(* IEC 61131-3 sources: virtual-bottling-plant/plc/src/process, 4 files *)

(* ---- FB_MixBatch.st ---- *)
(* T-101 batch sequence (PLC-03, ISA-88 phases): Fill (dose water, concentrate, sugar by
   flow totals), Mix, Transfer to T-301 through P-201. A recipe with another product first
   drains T-101 and T-301, then runs CIP. There is no time-of-day window: a new batch starts
   whenever T-101 is empty. One mix tank only (decision P2, see l1-plc.md). *)
FUNCTION_BLOCK FB_MixBatch
  VAR_INPUT
    Recipe : ST_Recipe;
    WaterFlow : REAL;        (* FT101, L/min *)
    ConcFlow : REAL;         (* FT102 *)
    SugarFlow : REAL;        (* FT103 *)
    Brix : REAL;             (* AT101 *)
    TankEmpty : BOOL;        (* LSL101 *)
    BufferLevel : REAL;      (* LT301, % *)
    CipDone : BOOL;
    NowMs : UDINT;
    DtS : REAL;
  END_VAR
  VAR_OUTPUT
    WaterValve : BOOL;
    ConcValve : BOOL;
    SugarValve : BOOL;
    Agitator : BOOL;
    TransferPump : BOOL;
    TankDrain : BOOL;
    BufferDrain : BOOL;
    CipRun : BOOL;
    ConcSelect : REAL;       (* product code to the concentrate feed selector *)
    Status : ST_T101Status;
    BrixAlarm : BOOL;
  END_VAR
  VAR
    MixTimer : FB_SimTon;
    NotEmptyInIdle : FB_SimTon;
    TargetWater : REAL;
    TargetConc : REAL;
    TargetSugar : REAL;
    DosedWater : REAL;
    DosedConc : REAL;
    DosedSugar : REAL;
    ConcBrix : REAL;
    PumpOn : BOOL;
  END_VAR
  VAR CONSTANT
    BATCH_L : REAL := 5000.0;
    SUGAR_SYRUP_BRIX : REAL := 67.0;
    MIX_MS : UDINT := 900000;        (* 15 min *)
    BUFFER_PUMP_ON : REAL := 90.0;   (* % T-301 *)
    BUFFER_PUMP_OFF : REAL := 98.0;
    BUFFER_EMPTY : REAL := 0.5;
  END_VAR

  WaterValve := FALSE; ConcValve := FALSE; SugarValve := FALSE; Agitator := FALSE;
  TransferPump := FALSE; TankDrain := FALSE; BufferDrain := FALSE; CipRun := FALSE;
  IF Status.ProductCode = 0 THEN
    Status.ProductCode := Recipe.ProductCode;  (* cold start: assume the recipe's product *)
  END_IF;

  NotEmptyInIdle(IN := Status.Phase = PHASE_IDLE AND NOT TankEmpty, PT := 10000,
                 NowMs := NowMs);
  CASE Status.Phase OF
    PHASE_IDLE:
      IF Recipe.ProductCode <> Status.ProductCode THEN
        Status.Phase := PHASE_DRAIN;
      ELSIF TankEmpty THEN
        IF Status.ProductCode = 2 THEN ConcBrix := 70.0; ELSE ConcBrix := 65.0; END_IF;
        TargetConc := Recipe.ConcRatio * BATCH_L;
        TargetSugar := MAX(0.0, (Recipe.BrixTarget - Recipe.ConcRatio * ConcBrix) * BATCH_L
                                / SUGAR_SYRUP_BRIX);
        TargetWater := BATCH_L - TargetConc - TargetSugar;
        DosedWater := 0.0; DosedConc := 0.0; DosedSugar := 0.0;
        Status.BatchNo := (Status.BatchNo + 1) MOD 30000;
        Status.BatchActive := TRUE;
        Status.BrixOk := FALSE;
        Status.BatchBrix := 0.0;
        BrixAlarm := FALSE;
        Status.Phase := PHASE_FILL;
      ELSIF NotEmptyInIdle.Q THEN
        (* Content of unknown dosing, e.g. after a PLC restart mid-batch: mix it, check the
           Brix and transfer it as its own batch rather than wait forever for an empty tank.
           Debounced: a sim reset clears its registers, so LSL101 reads 'not empty' briefly. *)
        Status.BatchNo := (Status.BatchNo + 1) MOD 30000;
        Status.BatchActive := TRUE;
        Status.Phase := PHASE_MIX;
      END_IF;

    PHASE_FILL:
      DosedWater := DosedWater + WaterFlow * DtS / 60.0;
      DosedConc := DosedConc + ConcFlow * DtS / 60.0;
      DosedSugar := DosedSugar + SugarFlow * DtS / 60.0;
      WaterValve := DosedWater < TargetWater;
      ConcValve := DosedConc < TargetConc;
      SugarValve := DosedSugar < TargetSugar;
      IF NOT (WaterValve OR ConcValve OR SugarValve) THEN
        Status.Phase := PHASE_MIX;
      END_IF;

    PHASE_MIX:
      Agitator := TRUE;
      IF MixTimer.Q THEN
        Status.BatchBrix := Brix;
        Status.BrixOk := ABS(Brix - Recipe.BrixTarget) <= Recipe.BrixTol;
        BrixAlarm := NOT Status.BrixOk;
        PumpOn := FALSE;
        Status.Phase := PHASE_TRANSFER;
      END_IF;

    PHASE_TRANSFER:
      Agitator := TRUE;
      IF BufferLevel < BUFFER_PUMP_ON THEN
        PumpOn := TRUE;
      ELSIF BufferLevel > BUFFER_PUMP_OFF THEN
        PumpOn := FALSE;
      END_IF;
      TransferPump := PumpOn AND NOT TankEmpty;
      IF TankEmpty THEN
        Status.BatchActive := FALSE;
        Status.Phase := PHASE_IDLE;
      END_IF;

    PHASE_DRAIN:
      TankDrain := NOT TankEmpty;
      BufferDrain := BufferLevel >= BUFFER_EMPTY;
      IF TankEmpty AND BufferLevel < BUFFER_EMPTY THEN
        Status.BatchActive := FALSE;
        Status.Phase := PHASE_CIP;
      END_IF;

    PHASE_CIP:
      CipRun := NOT CipDone;
      IF CipDone THEN
        Status.ProductCode := Recipe.ProductCode;
        Status.Phase := PHASE_IDLE;
      END_IF;
  END_CASE;

  MixTimer(IN := Status.Phase = PHASE_MIX, PT := MIX_MS, NowMs := NowMs);
  ConcSelect := INT_TO_REAL(Status.ProductCode);
END_FUNCTION_BLOCK

(* ---- FB_Pasteurizer.st ---- *)
(* P-201 HTST pasteuriser (PLC-12): outlet temperature PI on the steam valve with flow
   feedforward, and the divert valve. Without feedforward a step from recirculation to
   transfer flow drops the outlet below 83 °C for minutes (Phase 1 finding).
   The temperature rise per % steam scales with 1 / flow (8x at recirculation), so the gain
   is scheduled on flow. On a pump start or stop the flow measurement arrives a poll cycle
   late; the feedforward uses the commanded flow until FT201 agrees with it.
   Divert (PLC-11): opens at once below 83 °C; closes after 30 s stable at SP - 0.5 °C or more. *)
FUNCTION_BLOCK FB_Pasteurizer
  VAR_INPUT
    OutTemp : REAL;          (* TT202, °C *)
    Flow : REAL;             (* FT201, L/min *)
    SteamPressure : REAL;    (* PT201, bar *)
    TempSPCmd : REAL;        (* engineering setpoint from the bridge, 0 = keep *)
    PumpCmd : BOOL;          (* P101 transfer pump commanded *)
    NowMs : UDINT;
    DtS : REAL;
  END_VAR
  VAR_OUTPUT
    SteamValve : REAL;       (* TCV201, % *)
    Divert : BOOL := TRUE;   (* XV203, fail-safe: divert until proven hot *)
    Status : ST_P201Status;
    LowTempAlarm : BOOL;
    SteamLowAlarm : BOOL;
  END_VAR
  VAR
    TempCtrl : FB_PID;
    StableHot : FB_SimTon;
    SteamLow : FB_SimTon;
    DivertEdge : R_TRIG;
    Setpoint : REAL := 85.0;
    ExpectedFlow : REAL;
    FlowFF : REAL;
  END_VAR
  VAR CONSTANT
    MIN_SAFE_TEMP : REAL := 83.0;
    STABLE_MS : UDINT := 30000;
    NOMINAL_FLOW : REAL := 400.0;   (* L/min transfer *)
    RECIRC_FLOW : REAL := 50.0;     (* L/min, pump off *)
    FF_AT_NOMINAL : REAL := 60.0;   (* % steam valve at nominal flow *)
    KP_AT_NOMINAL : REAL := 2.0;    (* % per °C at nominal flow *)
    TI_S : REAL := 60.0;
    STEAM_LOW_BAR : REAL := 2.4;    (* nominal 3.0 bar *)
  END_VAR

  IF TempSPCmd >= 70.0 AND TempSPCmd <= 90.0 THEN
    Setpoint := TempSPCmd;
  END_IF;

  IF PumpCmd THEN
    ExpectedFlow := NOMINAL_FLOW;
  ELSE
    ExpectedFlow := RECIRC_FLOW;
  END_IF;
  IF ABS(Flow - ExpectedFlow) > 0.2 * ExpectedFlow THEN
    FlowFF := ExpectedFlow;               (* pump just started or stopped *)
  ELSE
    FlowFF := MAX(Flow, RECIRC_FLOW);
  END_IF;
  TempCtrl(Enable := TRUE, PV := OutTemp, SP := Setpoint,
           FF := FF_AT_NOMINAL * FlowFF / NOMINAL_FLOW,
           Kp := KP_AT_NOMINAL * FlowFF / NOMINAL_FLOW, Ti_s := TI_S, Td_s := 0.0,
           DtS := DtS, OutMin := 0.0, OutMax := 100.0);
  SteamValve := TempCtrl.Out;

  StableHot(IN := OutTemp >= Setpoint - 0.5, PT := STABLE_MS, NowMs := NowMs);
  IF OutTemp < MIN_SAFE_TEMP THEN
    Divert := TRUE;
  ELSIF StableHot.Q THEN
    Divert := FALSE;
  END_IF;
  DivertEdge(CLK := Divert);
  IF DivertEdge.Q THEN
    Status.DivertCount := (Status.DivertCount + 1) MOD 30000;
  END_IF;

  SteamLow(IN := SteamPressure < STEAM_LOW_BAR, PT := 5000, NowMs := NowMs);
  LowTempAlarm := OutTemp < MIN_SAFE_TEMP;
  SteamLowAlarm := SteamLow.Q;
  Status.TempSP := Setpoint;
  Status.ForwardFlowOk := NOT Divert;
END_FUNCTION_BLOCK

(* ---- FB_PID.st ---- *)
(* PI(D) controller with feedforward and anti-windup by conditional integration: the integral
   only moves when the output is not saturated in the direction the error pushes it.
   Dt comes from the sim clock (PLC-14), so tuning holds under time acceleration. *)
FUNCTION_BLOCK FB_PID
  VAR_INPUT
    Enable : BOOL;
    PV : REAL;
    SP : REAL;
    FF : REAL;          (* feedforward, added to the output *)
    Kp : REAL;          (* output % per unit of error *)
    Ti_s : REAL;        (* integral time, s (0 = no integral) *)
    Td_s : REAL;        (* derivative time on PV, s *)
    DtS : REAL;
    OutMin : REAL;
    OutMax : REAL;
  END_VAR
  VAR_OUTPUT
    Out : REAL;
    Error : REAL;
  END_VAR
  VAR
    ITerm : REAL;
    NextITerm : REAL;
    Unclamped : REAL;
    LastPV : REAL;
    DTerm : REAL;
  END_VAR

  Error := SP - PV;
  IF NOT Enable THEN
    ITerm := 0.0;
    Out := OutMin;
  ELSE
    IF DtS > 0.0 THEN
      DTerm := -Kp * Td_s * (PV - LastPV) / DtS;
      IF Ti_s > 0.0 THEN
        NextITerm := ITerm + Kp * Error * DtS / Ti_s;
        Unclamped := FF + Kp * Error + NextITerm + DTerm;
        IF (Unclamped < OutMax OR Error < 0.0) AND (Unclamped > OutMin OR Error > 0.0) THEN
          ITerm := NextITerm;
        END_IF;
      END_IF;
    END_IF;
    Out := LIMIT(OutMin, FF + Kp * Error + ITerm + DTerm, OutMax);
  END_IF;
  LastPV := PV;
END_FUNCTION_BLOCK

(* ---- FB_Tank.st ---- *)
(* Tank level monitor with a low-level hysteresis (T-301 filler interlock, PLC-11):
   Low below LowLimit, clears only at or above LowReset. *)
FUNCTION_BLOCK FB_Tank
  VAR_INPUT
    Level : REAL;        (* % *)
    LowLimit : REAL;     (* % *)
    LowReset : REAL;     (* % *)
  END_VAR
  VAR_OUTPUT
    Low : BOOL := TRUE;
    AboveLow : BOOL;
  END_VAR

  IF Level < LowLimit THEN
    Low := TRUE;
  ELSIF Level >= LowReset THEN
    Low := FALSE;
  END_IF;
  AboveLow := NOT Low;
END_FUNCTION_BLOCK
